Fanuc KAREL source: KT00907.KL

PROGRAM KT00907
%NOLOCKGROUP
%ENVIRONMENT VECTR
VAR
  V1: VECTOR
  V2: VECTOR
  OUT: VECTOR
BEGIN
  V1.X = 1.0
  V2.Y = 2.0
  V1.X = 1.0
  V2.Y = 2.0
  OUT = APPROACH(V1)
END KT00907
